(* PLC project Vn_tof_call, Beckhoff Automation GmbH TwinCAT PLC Control 3.5.13.21 *)
(* stored: creationDateTime 1970-01-01T00:00:00 *)

PROGRAM Vn_tof_call

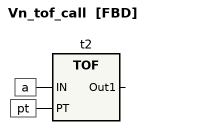
(* FBD diagram, written out as Structured Text *)
t2(IN := a, PT := pt);
END_PROGRAM
